(* IEC 61131-3 sources: SRCI_CLIENT_PLC/RobotLibrary/Library/POUs/General/MC_RobotTask (part 5) *)

           // Create log entry
           CreateLogMessagePara3 ( Timestamp   := SystemTime,
                                   MessageType := MessageType.CMD,
                                   Severity    := Severity.DEBUG,
                                   MessageCode := 0,
                                   MessageText := 'SyncWorkArea: Synchronization of WorkArea[{1}] triggered by PLC, SyncMode = {2}, SyncTime = {3}, SyncDirection = RC -> PLC',
                                   Para1       :=  DINT_TO_STRING(_rSyncIdx),
                                   Para2       :=  SYNC_MODE_TO_STRING(AxesGroup.Parameter.Plc.Parameter.SynchronizationModes.WorkAreas[SyncTime.AFTER_START_UP]),
                                   Para3       :=  SYNC_TIME_TO_STRING(SyncTime.AFTER_START_UP));
                                   RETURN;
         END_IF

         // Conflict triggered by RC ?
         IF ( NOT AxesGroup.State.SyncStateRc.InSync.WorkArea )
         THEN
           // get changed index
          _rSyncIdx := LIMIT(0, AxesGroup.State.SyncStateRc.UnSyncNo.WorkArea, AxesGroup.State.UnifiedWorkAreaIndex);
           // set timeout
           SetTimeout(PT := _rTimeout, rTimer := _rTimer);
           // inc step counter
          _rStep := 20; // -> read RC data and write it to PLC

           // Create log entry
           CreateLogMessagePara3 ( Timestamp   := SystemTime,
                                   MessageType := MessageType.CMD,
                                   Severity    := Severity.DEBUG,
                                   MessageCode := 0,
                                   MessageText := 'SyncWorkArea: Synchronization of WorkArea[{1}] triggered by RC, SyncMode = {2}, SyncTime = {3}, SyncDirection = RC -> PLC',
                                   Para1       :=  DINT_TO_STRING(_rSyncIdx),
                                   Para2       :=  SYNC_MODE_TO_STRING(AxesGroup.Parameter.Plc.Parameter.SynchronizationModes.WorkAreas[SyncTime.AFTER_START_UP]),
                                   Para3       :=  SYNC_TIME_TO_STRING(SyncTime.AFTER_START_UP));
                                   RETURN;
  			 END_IF

         // set timeout
         SetTimeout(PT := _rTimeout, rTimer := _rTimer);
         // jump back
        _rStep := 10;

    // ------------------------------------------
    // SyncMode : AUTOMATIC
    // ------------------------------------------
    13 : // Conflict triggerd by PLC ?
         IF ( NOT AxesGroup.State.SyncStatePlc.InSync.WorkArea )
         THEN
           // search for changed index
           FOR _rSyncIdx := 0 TO AxesGroup.State.UnifiedWorkAreaIndex
           DO
             IF ( AxesGroup.State.DataChanged.WorkArea[_rSyncIdx] )
             THEN
               // set timeout
               SetTimeout(PT := _rTimeout, rTimer := _rTimer);
               // inc step counter
              _rStep := 30; // -> write PLC data to RC
               EXIT;
  					 END_IF
           END_FOR

           // Create log entry
           CreateLogMessagePara3 ( Timestamp   := SystemTime,
                                   MessageType := MessageType.CMD,
                                   Severity    := Severity.DEBUG,
                                   MessageCode := 0,
                                   MessageText := 'SyncWorkArea: Synchronization of WorkArea[{1}] triggered by PLC, SyncMode = {2}, SyncTime = {3}, SyncDirection = PLC -> RC',
                                   Para1       :=  DINT_TO_STRING(_rSyncIdx),
                                   Para2       :=  SYNC_MODE_TO_STRING(AxesGroup.Parameter.Plc.Parameter.SynchronizationModes.WorkAreas[SyncTime.AFTER_START_UP]),
                                   Para3       :=  SYNC_TIME_TO_STRING(SyncTime.AFTER_START_UP));
                                   RETURN;
         END_IF

         // Conflict triggered by RC ?
         IF ( NOT AxesGroup.State.SyncStateRc.InSync.WorkArea )
         THEN
           // get changed index
          _rSyncIdx := LIMIT(0, AxesGroup.State.SyncStateRc.UnSyncNo.WorkArea, AxesGroup.State.UnifiedWorkAreaIndex);
           // set timeout
           SetTimeout(PT := _rTimeout, rTimer := _rTimer);
           // inc step counter
          _rStep := 20; // -> read RC data an write it to PLC

           // Create log entry
           CreateLogMessagePara3 ( Timestamp   := SystemTime,
                                   MessageType := MessageType.CMD,
                                   Severity    := Severity.DEBUG,
                                   MessageCode := 0,
                                   MessageText := 'SyncWorkArea: Synchronization of WorkArea[{1}] triggered by RC, SyncMode = {2}, SyncTime = {3}, SyncDirection = RC -> PLC',
                                   Para1       :=  DINT_TO_STRING(_rSyncIdx),
                                   Para2       :=  SYNC_MODE_TO_STRING(AxesGroup.Parameter.Plc.Parameter.SynchronizationModes.WorkAreas[SyncTime.AFTER_START_UP]),
                                   Para3       :=  SYNC_TIME_TO_STRING(SyncTime.AFTER_START_UP));
                                   RETURN;
  			 END_IF

         // set timeout
         SetTimeout(PT := _rTimeout, rTimer := _rTimer);
         // jump back
        _rStep := 10; // ST-FIX F95: was commented out

    // ------------------------------------------
    // Read Data from RC and write it to PLC
    // ------------------------------------------
    20 : IF (( NOT _readWorkArea.Busy  ) AND
             ( NOT _readWorkArea.Error ))
         THEN
           // set command parameter
          _readWorkArea.ParCmd.WorkAreaNo := _rSyncIdx;
           // execute command
          _readWorkArea.Execute := TRUE;
           // set timeout
           SetTimeout(PT := _rTimeout, rTimer := _rTimer);
           // inc step counter
          _rStep := _rStep + 1;
         ELSE
           // check error ?
           IF (_readWorkArea.Error)
           THEN
             ErrorID     := _readWorkArea.ErrorID;
             ErrorAddTxt := _readWorkArea.ErrorAddTxt;
           END_IF

           // timeout exceeded ?
           IF (CheckTimeout(_rTimer) = RobotLibraryConstants.OK)
           THEN
             ErrorID     := RobotLibraryErrorIdEnum.ERR_TIMEOUT_CMD;
             ErrorAddTxt := CONCAT(_stepName, DINT_TO_STRING(_rStep));
           END_IF
         END_IF

    21 : IF (( NOT _readWorkArea.Busy  ) AND
             ( NOT _readWorkArea.Error ) AND
             (     _readWorkArea.Done  ))
         THEN
           // reset execution
          _readWorkArea.Execute := FALSE;
           // ST-FIX F107: AUTOMATIC - the PLC data were changed while the RC data were read: the PLC
           // change is the most recent one and is written to the RC instead of being overwritten
           IF ( AxesGroup.Parameter.Plc.Parameter.SynchronizationModes.WorkAreas[SyncTime.AFTER_START_UP] = SyncMode.AUTOMATIC ) AND
              ( NOT IsWorkAreaEqual( Data1 := WorkAreas[_rSyncIdx].Data, Data2 := _workAreas[_rSyncIdx].Data, IgnoreTimestamp := TRUE ))
           THEN
             // set timeout
             SetTimeout(PT := _rTimeout, rTimer := _rTimer);
             // -> write PLC data to RC
            _rStep := 30;
             RETURN;
           END_IF
           // update internal WorkArea data
           WorkAreas[_rSyncIdx].Data := _readWorkArea.OutCmd.WorkAreaData;
          _workAreas[_rSyncIdx].Data := _readWorkArea.OutCmd.WorkAreaData;
           // set available bit
           WorkAreas[_rSyncIdx].Available := TRUE;
          _workAreas[_rSyncIdx].Available := TRUE;
           // set timeout
           SetTimeout(PT := _rTimeout, rTimer := _rTimer);
           // inc step counter
          // ST-FIX F20: write the RC data back to reset DataChanged on the RC (spec 5.6.7.4.2)
          IF ( AxesGroup.State.RobotData.RCSupportedFunctions.WriteWorkArea )
          THEN
            _rStep := 30;
          ELSE
            _rStep := 10;
          END_IF // -> jump to after startup
         ELSE
           // check error ?
           IF (_readWorkArea.Error)
           THEN
             ErrorID     := _readWorkArea.ErrorID;
             ErrorAddTxt := _readWorkArea.ErrorAddTxt;
             // reset available bit
             WorkAreas[_rSyncIdx].Available := FALSE;
            _workAreas[_rSyncIdx].Available := FALSE;
           END_IF

           // timeout exceeded ?
           IF (CheckTimeout(_rTimer) = RobotLibraryConstants.OK)
           THEN
             ErrorID     := RobotLibraryErrorIdEnum.ERR_TIMEOUT_CMD;
             ErrorAddTxt := CONCAT(_stepName, DINT_TO_STRING(_rStep));
           END_IF
         END_IF

    // ------------------------------------------
    // Write data from PLC to RC
    // ------------------------------------------
    30 : IF (( NOT _writeWorkArea.Busy  ) AND
             ( NOT _writeWorkArea.Error ))
         THEN
           // set command parameter
          _writeWorkArea.ParCmd.WorkAreaNo   := _rSyncIdx;
          _writeWorkArea.ParCmd.WorkAreaData :=  WorkAreas[_rSyncIdx].Data;
           // execute command
          _writeWorkArea.Execute := TRUE;
           // set timeout
           SetTimeout(PT := _rTimeout, rTimer := _rTimer);
           // inc step counter
          _rStep := _rStep + 1;
         ELSE
           // check error ?
           IF (_writeWorkArea.Error)
           THEN
             ErrorID     := _writeWorkArea.ErrorID;
             ErrorAddTxt := _writeWorkArea.ErrorAddTxt;;
           END_IF

           // timeout exceeded ?
           IF (CheckTimeout(_rTimer) = RobotLibraryConstants.OK)
           THEN
             ErrorID     := RobotLibraryErrorIdEnum.ERR_TIMEOUT_CMD;
             ErrorAddTxt := CONCAT(_stepName, DINT_TO_STRING(_rStep));
           END_IF
         END_IF

    31 : IF (( NOT _writeWorkArea.Busy  ) AND
             ( NOT _writeWorkArea.Error ) AND
             (     _writeWorkArea.Done  ))
         THEN
           // execute command
          _writeWorkArea.Execute := FALSE;
           // update internal WorkArea data
          _workAreas[_rSyncIdx] := WorkAreas[_rSyncIdx];
           // set available bit
           WorkAreas[_rSyncIdx].Available := TRUE;
          _workAreas[_rSyncIdx].Available := TRUE;
           // set timeout
           SetTimeout(PT := _rTimeout, rTimer := _rTimer);
           // inc step counter
          _rStep := 10; // -> jump to after startup;
         ELSE
           // check error ?
           IF (_writeWorkArea.Error)
           THEN
             SetWarning( WarningID := RobotLibraryWarningIdEnum.WARN_WORK_AREA_SYNC_FAILED_BY_ERROR_OF_READ_OR_WRITE_CMD, Overwrite :=  TRUE);
             // reset available bit
             WorkAreas[_rSyncIdx].Available := FALSE;
            _workAreas[_rSyncIdx].Available := FALSE;
           END_IF

           // timeout exceeded ?
           IF (CheckTimeout(_rTimer) = RobotLibraryConstants.OK)
           THEN
             ErrorID     := RobotLibraryErrorIdEnum.ERR_TIMEOUT_CMD;
             ErrorAddTxt := CONCAT(_stepName, DINT_TO_STRING(_rStep));
           END_IF
         END_IF

  ELSE
    // invalid step
    ErrorID     := RobotLibraryErrorIdEnum.ERR_INVALID_STEP;
    ErrorAddTxt := CONCAT(_stepName , DINT_TO_STRING(_stepCmd));
  END_CASE

END_METHOD

METHOD PRIVATE HandleTelegramStateCtrl
VAR_INPUT
END_VAR

  // Telegram Control
  // ----------------
  IF ( _lastTelegramControl <> GetHalfeByteLo(Telegram.PlcToRob.Header.AxesGroupID_Control))
  THEN
    // Create log entry
    CreateLogMessagePara2 ( Timestamp   := SystemTime,
                            MessageType := MessageType.CMD,
                            Severity    := Severity.INFO,
                            MessageCode := 0,
                            MessageText := 'SRCI Interface control changed from {1} to {2}',
                            Para1       := TELEGRAM_CONTROL_TO_STRING(_lastTelegramControl),
                            Para2       := TELEGRAM_CONTROL_TO_STRING(GetHalfeByteLo(Telegram.PlcToRob.Header.AxesGroupID_Control)));

    _lastTelegramControl := GetHalfeByteLo(Telegram.PlcToRob.Header.AxesGroupID_Control);
  END_IF

  // Telegram State
  // ----------------
  IF ( _lastTelegramState <> Telegram.RobToPlc.Header.TelegramState)
  THEN
    // Create log entry
    CreateLogMessagePara2 ( Timestamp   := SystemTime,
                            MessageType := MessageType.CMD,
                            Severity    := Severity.INFO,
                            MessageCode := 0,
                            MessageText := 'SRCI Interface state changed from {1} to {2}',
                            Para1       := TELEGRAM_STATE_TO_STRING(_lastTelegramState),
                            Para2       := TELEGRAM_STATE_TO_STRING(Telegram.RobToPlc.Header.TelegramState));

    // Check Interface changed after being initialized ?
    IF ((  Enable                                                                          ) AND
        ( _lastTelegramState                      = TelegramState.INITIALIZED              ) AND
       ((  Telegram.RobToPlc.Header.TelegramState = TelegramState.READY_FOR_INITIALIZATION ) OR
        (  Telegram.RobToPlc.Header.TelegramState = TelegramState.READY_TO_RESUME          )))
    THEN
      // the error 16#80A7 (interface reset after the initialization) is set in OnCall (ST-FIX F65)
      ;
  	END_IF

    // apply new telegram state
   _lastTelegramState := Telegram.RobToPlc.Header.TelegramState;
  END_IF

END_METHOD

METHOD HandleUserData
VAR_IN_OUT
   /// Robot assignment of function
  AxesGroup    : AxesGroup;
  ///  User data stored on the PLC according to Table 6-10
  UserData     : UserData;
END_VAR

  // Common
  UserData.LogLevel                          := LogLevel;

  UserData.PLCManufacturedID                 := _parCfg.Plc.Parameter.ManufacturedID;
  UserData.PLCOrderID                        := _parCfg.Plc.Parameter.OrderID;
  UserData.PLCSerialNumber                   := _parCfg.Plc.Parameter.SerialNumber;
  UserData.PLCFirmwareVersion                := _parCfg.Plc.Parameter.FirmwareVersion;
  UserData.PLCInterfaceVersion               := _parCfg.Plc.Parameter.InterfaceVersion;
  UserData.PLCLibraryVersion                 :=  RobotLibraryConstants.PLCLibraryVersion;

  // Communication
  UserData.LifeSignTimeOut                   := _parCfg.Com.LifeSignTimeOut;

  // Plc Parameter
  UserData.SynchronizationModes              := _parCfg.Plc.Parameter.SynchronizationModes;
  UserData.EnableSync                        :=  SyncModesToDataEnableSync(Value := _parCfg.Plc.Parameter.SynchronizationModes);

  // Robot Parameter
  UserData.DelayTime                         := _parCfg.Rob.Parameter.DelayTime;
  UserData.WaitForNrOfCmd                    := _parCfg.Rob.Parameter.WaitForNrOfCmd;
  UserData.WaitAtBlendingZone                := _parCfg.Rob.Parameter.WaitAtBlendingZone;
  UserData.AllowSecSeqWhileSubprogram        := _parCfg.Rob.Parameter.AllowSecSeqWhileSubprogram;
  UserData.AllowDynamicBlending              := _parCfg.Rob.Parameter.AllowDynamicBlending;
  UserData.SyncReaction                      := _parCfg.Rob.Parameter.SyncReaction;
  UserData.SyncDelay                         := _parCfg.Rob.Parameter.SyncDelay;
  UserData.MessageLevel                      := _parcfg.Rob.Parameter.MessageLevel;

  // ReadRobotData
  UserData.RCManufacturer                    := AxesGroup.State.RobotData.RCManufacturer;
  UserData.RCOrderID                         := AxesGroup.State.RobotData.RCOrderID;
  UserData.RCSerialNumber                    := AxesGroup.State.RobotData.RCSerialNumber;
  UserData.RASerialNumber                    := AxesGroup.State.RobotData.RASerialNumber;
  UserData.RCFirmwareVersion                 := AxesGroup.State.RobotData.RCFirmwareVersion;

  UserData.RCInterpreterVersion := AxesGroup.State.RobotData.RCInterpreterVersionNumber; // ST-FIX F163: was characters 1/2/3 of the text

  UserData.AxisJointUsed                     := AxesGroup.State.RobotData.AxisJointUsed;
  UserData.AxisExternalUsed                  := AxesGroup.State.RobotData.AxisExternalUsed;
  UserData.AxisJointUnit                     := AxesGroup.State.RobotData.AxisJointUnit;
  UserData.AxisExternalUnit                  := AxesGroup.State.RobotData.AxisExternalUnit;
  UserData.RCSupportedFunctions              := AxesGroup.State.RobotData.RCSupportedFunctions;

  UserData.BrakeTestRequired                 := AxesGroup.State.ConfigurationData.BrakeTestRequired;
  UserData.PathAccuracyMode                  := AxesGroup.State.ConfigurationData.PathAccuracyMode;
  UserData.AvoidSingularity                  := AxesGroup.State.ConfigurationData.AvoidSingularity;
  UserData.ConstantVelocitySupported         := AxesGroup.State.ConfigurationData.ConstantVelocitySupported;
  UserData.StepModeExactStopActive           := AxesGroup.State.ConfigurationData.StepModeExactStopActive;
  UserData.StepModeBlendingActive            := AxesGroup.State.ConfigurationData.StepModeBlendingActive;
  UserData.AcceleratingSupported             := AxesGroup.State.ConfigurationData.AcceleratingSupported;
  UserData.DeceleratingSupported             := AxesGroup.State.ConfigurationData.DecceleratingSupported;

  UserData.Initialized                       := Initialized;
  UserData.Synchronized                      := Synchronized;

  // Cyclic data
  UserData.RCSRCIVersion                     := AxesGroup.Cyclic.RobToPlc.SRCIVersion;
  UserData.IsMoving                          := AxesGroup.Cyclic.RobToPlc.StatusRobotArm.IsMoving;
  UserData.PrimarySequencePaused             := AxesGroup.Cyclic.RobToPlc.StatusRobotArm.PrimarySequencePaused;
  UserData.InPrimaryPos                      := AxesGroup.Cyclic.RobToPlc.StatusRobotArm.InPrimaryPos;
  UserData.SecondarySequenceActive           := AxesGroup.Cyclic.RobToPlc.StatusRobotArm.SecondarySequenceActive;
  UserData.ErrorPending                      := AxesGroup.Cyclic.RobToPlc.StatusRobotArm.ErrorPending;
  UserData.RestartInProgress                 := AxesGroup.Cyclic.RobToPlc.StatusRobotArm.RestartInProgress;
  UserData.Enabled                           := AxesGroup.Cyclic.RobToPlc.StatusRobotArm.Enabled;
  UserData.Idle                              := AxesGroup.Cyclic.RobToPlc.StatusRobotArm.RaSequenceState = RaSequenceState.IDLE;
  UserData.Executing                         := AxesGroup.Cyclic.RobToPlc.StatusRobotArm.RaSequenceState = RaSequenceState.EXECUTING;
  UserData.Interrupted                       := AxesGroup.Cyclic.RobToPlc.StatusRobotArm.RaSequenceState = RaSequenceState.INTERRUPTED;
  UserData.IsBlending                        := AxesGroup.Cyclic.RobToPlc.StatusRobotArm.IsBlending;
  UserData.OperationMode                     := AxesGroup.Cyclic.RobToPlc.StatusRobotArm.OperationMode;
  UserData.CollisionDetectionEnabled         := AxesGroup.Parameter.Rob.Parameter.CollisionDetectionEnabled; // ST-FIX F169: the status word bit is always FALSE
  UserData.CollisionDetected                 := AxesGroup.Cyclic.RobToPlc.StatusRobotArm.CollisionDetected;
  UserData.RestartRequested                  := AxesGroup.Cyclic.RobToPlc.StatusRobotArm.RestartRequested;
  UserData.Accelerating                      := AxesGroup.Cyclic.RobToPlc.StatusRobotArm.Accelerating;
  UserData.Decelerating                      := AxesGroup.Cyclic.RobToPlc.StatusRobotArm.Decelerating;
  UserData.ConstantVelocity                  := AxesGroup.Cyclic.RobToPlc.StatusRobotArm.ConstantVelocity;
  UserData.ActualOverride                    := PERCENT_UINT_TO_REAL( Value := AxesGroup.Cyclic.RobToPlc.Override, IsOptional := FALSE);

  // Cyclic optional data
  UserData.CartesianPosition                 := AxesGroup.CyclicOptional.RobToPlc.CartesianPosition;
  UserData.ExtCartesianPosition              := AxesGroup.CyclicOptional.RobToPlc.CartesianPositionExt;
  UserData.JointPosition                     := AxesGroup.CyclicOptional.RobToPlc.JointPosition;
  UserData.ExtJointPosition                  := AxesGroup.CyclicOptional.RobToPlc.JointPositionExt;

  // Synchronizing
  UserData.ToolDataSynchronizing             := AxesGroup.State.Synchronizing.Tool;
  UserData.FrameDataSynchronizing            := AxesGroup.State.Synchronizing.Frame;
  UserData.LoadDataSynchronizing             := AxesGroup.State.Synchronizing.Load;
  UserData.WorkAreaDataSynchronizing         := AxesGroup.State.Synchronizing.WorkAreas;
  UserData.SWLimitsSynchronizing             := AxesGroup.State.Synchronizing.SwLimits;
  UserData.DefaultDynamicsSynchronizing      := AxesGroup.State.Synchronizing.DefaultDynamics;
  UserData.ReferenceDynamicsSynchronizing    := AxesGroup.State.Synchronizing.ReferenceDynamics;

  UserData.ActivateTwoSequences              := _parCfg.Com.TwoSequences;
  UserData.ReadingCartesianPosition          :=  AxesGroup.State.ReadingCartesianPosition;
  UserData.ReadingExtCartesianPosition       :=  AxesGroup.State.ReadingCartesianPositionExt;
  UserData.ReadingJointPosition              :=  AxesGroup.State.ReadingJointPosition;
  UserData.ReadingExtJointPosition           :=  AxesGroup.State.ReadingJointPositionExt;

END_METHOD

PROPERTY PROTECTED HasError : Bool

GET
VAR
END_VAR

  HasError := ErrorID <> RobotLibraryErrorIdEnum.NO_ERROR;

END_GET

PROPERTY PROTECTED HasInfo : BOOL

GET
VAR
END_VAR

  HasInfo := InfoID <> RobotLibraryInfoIdEnum.NO_INFO;

END_GET

PROPERTY PROTECTED HasWarning : BOOL

GET
VAR
END_VAR

  HasWarning := WarningID <> RobotLibraryWarningIdEnum.NO_WARNING;

END_GET

METHOD PRIVATE OnCall
VAR_IN_OUT
   /// Robot assignment of function
  AxesGroup : AxesGroup;
END_VAR

  // map numeric value to enum, so that the corresponding message text is directly shown by the tooltip
  ErrorIdEnum   := ErrorId;
  WarningIdEnum := WarningId;
  InfoIdEnum    := InfoId;

  Error := HasError;

  // Check Payload and In/Out data size
  IF (( ROBOT_IN_DATA_SIZE  < 64 ) OR
      ( ROBOT_OUT_DATA_SIZE < 64 ))
  THEN
    SetError(ErrorID := RobotLibraryErrorIdEnum.ERR_INVALID_LIBRARY_PARA, Overwrite := TRUE );
    RETURN;
  END_IF

  // Check AxesGroupID valid
  IF (( AxesGroupID < RobotLibraryConstants.AXES_GROUP_ID_MIN ) OR
      ( AxesGroupID > RobotLibraryConstants.AXES_GROUP_ID_MAX ))
  THEN
    // ST-FIX F138: client error of the specification (16#80AA, table 7-2) instead of the internal ID 3
    SetError( ErrorID := RobotLibraryErrorIdEnum.ERR_AXESGROUP_ID_INVALID_0x80AA, Overwrite := TRUE );
    RETURN;
  END_IF

  // Reset flag for initialization / Synchronization
  IF ( Initialized OR Synchronized) AND ( AxesGroup.Cyclic.RobToPlc.TelegramState <> TelegramState.INITIALIZED)
  THEN
    // Reset initialized flag
    Initialized := FALSE;
    // Reset Synchronized flag
    Synchronized := FALSE;
    // Set error
    // ST-FIX F65: reason of the loss of the initialization (table 7-2): RI error of the RC in the
    // telegram state (16#A1..16#AD), interface reset by the RC (16#80A7) or unknown (16#80A2)
    IF (( AxesGroup.Cyclic.RobToPlc.TelegramState >= TelegramState.ERROR_161_TELEGRAM_CONTROL_MISMATCH_TELEGRAM_STATE ) AND
        ( AxesGroup.Cyclic.RobToPlc.TelegramState <= TelegramState.ERROR_173_SERVER_CONNECTION_LOST                   ))
    THEN
      SetError( ErrorID := AxesGroup.Cyclic.RobToPlc.TelegramState, Overwrite := TRUE );
      // Create log entry
      CreateLogMessagePara1 ( Timestamp   := SystemTime,
                              MessageType := MessageType.CMD,
                              Severity    := Severity.ERROR,
                              MessageCode := ErrorID,
                              MessageText := 'Initialization lost: RI error {1} of the RC',
                              Para1       := TELEGRAM_STATE_TO_STRING(AxesGroup.Cyclic.RobToPlc.TelegramState));
    ELSIF (( AxesGroup.Cyclic.RobToPlc.TelegramState = TelegramState.READY_FOR_INITIALIZATION ) OR
           ( AxesGroup.Cyclic.RobToPlc.TelegramState = TelegramState.READY_TO_RESUME          ))
    THEN
      SetError( ErrorID := RobotLibraryErrorIdEnum.ERR_INTERFACE_WAS_RESET_AFTER_INIT_0x80A7, Overwrite := TRUE );
      // Create log entry
      CreateLogMessagePara1 ( Timestamp   := SystemTime,
                              MessageType := MessageType.CMD,
                              Severity    := Severity.ERROR,
                              MessageCode := ErrorID,
                              MessageText := 'Initialization lost: interface was reset by the RC (state {1})',
                              Para1       := TELEGRAM_STATE_TO_STRING(AxesGroup.Cyclic.RobToPlc.TelegramState));
    ELSE
      SetError( ErrorID := RobotLibraryErrorIdEnum.ERR_INIT_LOST_UNKNOWN_0x80A2, Overwrite := TRUE );
      // Create log entry
      CreateLogMessagePara1 ( Timestamp   := SystemTime,
                              MessageType := MessageType.CMD,
                              Severity    := Severity.ERROR,
                              MessageCode := ErrorID,
                              MessageText := 'Initialization lost: unknown reason (state {1})',
                              Para1       := TELEGRAM_STATE_TO_STRING(AxesGroup.Cyclic.RobToPlc.TelegramState));
    END_IF
  END_IF

  // Warning for ACR Registers running low
  IF ( AxesGroup.Acyclic.ActiveCommandRegister.CurrentAcrUsagePercent > RobotLibraryParameter.ACR_USAGE_WARNING_LIMIT )
  THEN
    SetWarning( WarningID := RobotLibraryWarningIdEnum.WARN_ACR_FREE_ENTRIES_LOW, Overwrite := TRUE);
  END_IF

  // Check ToolData boundary
  IF ( AxesGroup.SystemData.ToolDataMin  <> 0 )
  THEN
    SetWarning( WarningID := RobotLibraryWarningIdEnum.WARN_TOOL_DATA_ARRAY_NOT_START_AT_ZERO, Overwrite := FALSE );
  END_IF

  // Check FrameData boundary
  IF ( AxesGroup.SystemData.FrameDataMin <> 0 ) AND ( NOT HasWarning )
  THEN
    SetWarning( WarningID := RobotLibraryWarningIdEnum.WARN_FRAME_DATA_ARRAY_NOT_START_AT_ZERO, Overwrite := FALSE );
  END_IF

  // Check WorkAreas boundary
  IF ( AxesGroup.SystemData.WorkAreasMin <> 0 ) AND ( NOT HasWarning )
  THEN
    SetWarning( WarningID := RobotLibraryWarningIdEnum.WARN_FRAME_DATA_ARRAY_NOT_START_AT_ZERO, Overwrite := FALSE);
  END_IF

  // Check configuration parameter changed ?
  CheckParameterChanged(AxesGroup := AxesGroup);

END_METHOD

METHOD OnExecRun : DINT
VAR_IN_OUT
  /// Robot assignment of function
  AxesGroup         : AxesGroup;
END_VAR

  // building rising and falling edges
  _enable_R( CLK := Enable);
  _enable_F( CLK := Enable);

  IF ( _enable_F.Q)
  THEN
    Reset(AxesGroup := AxesGroup);
  END_IF

  OnExecRun := RobotLibraryConstants.RUNNING;

  CASE _stepCmd OF

    00:  IF ( _enable_R.Q )
         THEN
           // Create log entry
           CreateLogMessage ( Timestamp   := SystemTime,
                              MessageType := MessageType.CMD,
                              Severity    := Severity.INFO,
                              MessageCode := 0,
                              MessageText := 'Robot Task Enabled');

           // reset the rising edge
          _enable_R();
           // set busy flag
           Busy := TRUE;
           // set timeout
           SetTimeout(PT := _timeoutCmd, rTimer := _timerCmd);
           // Reset FastStop
           AxesGroup.Cyclic.PlcToRob.FastStop := 0;
           // Reset Active command register
           AxesGroup.Acyclic.ActiveCommandRegister.Reset();
           // ST-FIX F23: the RC is still initialized from the previous enable (ACR, SEQ/ACK)
           // -> reset the interface on the RC as well
           _restartReset := AxesGroup.Cyclic.RobToPlc.TelegramState = TelegramState.INITIALIZED;
           IF ( _restartReset )
           THEN
             AxesGroup.Cyclic.PlcToRob.Control := ControlHalfByte.RESET;
           END_IF

           // check parameter valid
           IF ( CheckParameterValid(AxesGroup := AxesGroup) )
           THEN
             // take configuration parameter if not yet enabled
            _parCfg := ParCfg;
            // ST-FIX F103: number of telegram sequences of this configuration (not of the previous enable)
            IF ( _parCfg.Com.TwoSequences )
            THEN
              AxesGroup.State.SequenceCountSend := 1;
            ELSE
              AxesGroup.State.SequenceCountSend := 0;
            END_IF
            // ST-FIX F79: no error state of the RC seen yet in this initialization
            _initErrorState := TelegramState.UNDEFINED;
             // inc step counter
            _stepCmd := _stepCmd + 1;
           END_IF
         END_IF

    01:  // ST-FIX F153: INITIALIZED without a request of this RobotTask: the RC is still
  // initialized from an earlier connection -> reset the interface on the RC first
  IF (( AxesGroup.Cyclic.RobToPlc.TelegramState = TelegramState.INITIALIZED ) AND
      ( AxesGroup.Cyclic.PlcToRob.Control       = ControlHalfByte.NONE      ) AND
      ( NOT _restartReset                                                   ))
  THEN
    AxesGroup.Cyclic.PlcToRob.Control := ControlHalfByte.RESET;
    _restartReset := TRUE;
  END_IF

  // ST-FIX F23: wait until the RC left the state INITIALIZED of the previous enable
  IF ( _restartReset )
  THEN
    IF ( AxesGroup.Cyclic.RobToPlc.TelegramState <> TelegramState.INITIALIZED )
    THEN
      _restartReset := FALSE;
    END_IF
  ELSE
  CASE AxesGroup.Cyclic.RobToPlc.TelegramState  OF

           TelegramState.UNDEFINED : ;

           TelegramState.ERROR_161_TELEGRAM_CONTROL_MISMATCH_TELEGRAM_STATE..TelegramState.ERROR_172_TELEGRAM_NUMBER_NOT_SUPPORTED:

             // ST-FIX F79: remember the error state for the init timeout
             _initErrorState := AxesGroup.Cyclic.RobToPlc.TelegramState;

             // clear error
             AxesGroup.Cyclic.PlcToRob.Control := ControlHalfByte.ACK_ERROR;
             AxesGroup.Cyclic.PlcToRob.Control := ControlHalfByte.RESET; // always a reset, so that on the robot side the ACR is reseted

           TelegramState.ERROR_173_SERVER_CONNECTION_LOST:

             // Reset interface including the ACR register on server side
             AxesGroup.Cyclic.PlcToRob.Control := ControlHalfByte.RESET;

           TelegramState.READY_TO_RESUME :

             // Resume
             AxesGroup.Cyclic.PlcToRob.Control := ControlHalfByte.RESUME;

           TelegramState.READY_FOR_INITIALIZATION:

             // Request initialization
             AxesGroup.Cyclic.PlcToRob.Control := ControlHalfByte.INITIALIZE;

           TelegramState.INITIALIZED:

             // Reset Telegram Control
             AxesGroup.Cyclic.PlcToRob.Control := ControlHalfByte.NONE;

             // Check SRCI Version is compatible ?
             IF ( AxesGroup.Cyclic.RobToPlc.SRCIVersion.MajorVersion = RobotLibraryConstants.SRCIVersion.MajorVersion )
             THEN
               // set timeout
               SetTimeout(PT := _timeoutCmd, rTimer := _timerCmd);
               // inc step counter
              _stepCmd := _stepCmd + 1;
             ELSE
               // set error
               ErrorID     := RobotLibraryErrorIdEnum.ERR_SRCI_MAJOR_VERSION_INCOMPATIBLE_0x80A4;
               ErrorAddTxt := CONCAT('_stepCmd = ' , DINT_TO_STRING(_stepCmd));
             END_IF

         ELSE
           // TelegrammState in error
           SetError( ErrorID := RobotLibraryErrorIdEnum.ERR_INIT_LOST_UNKNOWN_0x80A2, Overwrite := TRUE ); // ST-FIX F65: unknown state (16#A2 is the RI error of the RC)
             // Create log entry
             CreateLogMessagePara1 ( Timestamp   := SystemTime,
                                     MessageType := MessageType.CMD,
                                     Severity    := Severity.ERROR,
                                     MessageCode := ErrorID,
                                     MessageText := 'Initialization lost: unknown telegram state {1}',
                                     Para1       := TELEGRAM_STATE_TO_STRING(AxesGroup.Cyclic.RobToPlc.TelegramState));
           ErrorAddTxt := CONCAT('_stepCmd = ' , DINT_TO_STRING(_stepCmd));
         END_CASE
  END_IF

         // timeout exceeded ?
         IF (CheckTimeout(_timerCmd) = RobotLibraryConstants.OK)
         THEN
           // Check Telegram State error ?
           IF (( AxesGroup.Cyclic.RobToPlc.TelegramState >= TelegramState.ERROR_161_TELEGRAM_CONTROL_MISMATCH_TELEGRAM_STATE ) AND // ST-FIX F15
               ( AxesGroup.Cyclic.RobToPlc.TelegramState <= TelegramState.ERROR_173_SERVER_CONNECTION_LOST                   ))
           THEN
             ErrorID     := AxesGroup.Cyclic.RobToPlc.TelegramState;
             ErrorAddTxt := CONCAT('_stepCmd = ' , DINT_TO_STRING(_stepCmd));
           ELSIF ( _initErrorState <> TelegramState.UNDEFINED ) // ST-FIX F79: error state seen during the initialization
           THEN
             ErrorID     := _initErrorState;
             ErrorAddTxt := CONCAT('_stepCmd = ' , DINT_TO_STRING(_stepCmd));
           ELSE
             ErrorID     := RobotLibraryErrorIdEnum.ERR_TIMEOUT_CMD;
             ErrorAddTxt := CONCAT('_stepCmd = ' , DINT_TO_STRING(_stepCmd));
           END_IF
         END_IF

    02: IF (( NOT _readMessages.Busy  ) AND
            ( NOT _readMessages.Error ))
        THEN
          // start function block
         _readMessages.Enable := TRUE;
         _readMessages.ParCmd.MsgID := 0;
         _readMessages.ParCmd.MessageLevel := _parCfg.Rob.Parameter.MessageLevel;

          // set timeout
          SetTimeout(PT := _timeoutCmd, rTimer := _timerCmd);
          // inc step counter
         _stepCmd := _stepCmd + 1;
        ELSE
          // check error ?
          IF (_readMessages.Error)
          THEN
            ErrorID     := _readMessages.ErrorID;
            ErrorAddTxt := _readMessages.ErrorAddTxt;;
          END_IF
          // timeout exceeded ?
          IF (CheckTimeout(_timerCmd) = RobotLibraryConstants.OK)
          THEN
            ErrorID     := RobotLibraryErrorIdEnum.ERR_TIMEOUT_CMD;
            ErrorAddTxt := CONCAT('_stepCmd = ' , DINT_TO_STRING(_stepCmd));
          END_IF
        END_IF

    03: IF ((     _readMessages.Enabled ) AND
            ( NOT _readMessages.Error   ))
        THEN
          // ---------------------------------------------------------------
          // !!! ReadMessages must stay active for the Message mechanism !!!
          // ---------------------------------------------------------------
          // ReadMessages.Enable := FALSE;
          // set timeout
          SetTimeout(PT := _timeoutCmd, rTimer := _timerCmd);
          // inc step counter
         _stepCmd := _stepCmd + 1;
        ELSE
           // check error ?
           IF (_readMessages.Error)
           THEN
             ErrorID     := _readMessages.ErrorID;
             ErrorAddTxt := _readMessages.ErrorAddTxt;;
           END_IF

           // timeout exceeded ?
           IF (CheckTimeout(_timerCmd) = RobotLibraryConstants.OK)
           THEN
             ErrorID     := RobotLibraryErrorIdEnum.ERR_TIMEOUT_CMD;
             ErrorAddTxt := CONCAT('_stepCmd = ' , DINT_TO_STRING(_stepCmd));
           END_IF
         END_IF

    04: IF (( NOT _exchangeConfiguration.Busy  ) AND
            ( NOT _exchangeConfiguration.Error ))
        THEN
          // set command parameter
         _exchangeConfiguration.ParCmd.LogLevel                           :=  LogLevel;
         _exchangeConfiguration.ParCmd.WaitAtBlendingZone                 := _parCfg.Rob.Parameter.WaitAtBlendingZone;
         _exchangeConfiguration.ParCmd.AllowSecSeqWhileSubprogram         := _parCfg.Rob.Parameter.AllowSecSeqWhileSubprogram;
         _exchangeConfiguration.ParCmd.AllowDynamicBlending               := _parCfg.Rob.Parameter.AllowDynamicBlending;
         _exchangeConfiguration.ParCmd.DelayTime                          := _parCfg.Rob.Parameter.DelayTime;
         _exchangeConfiguration.ParCmd.WaitForNrOfCmd                     := _parCfg.Rob.Parameter.WaitForNrOfCmd;
         _exchangeConfiguration.ParCmd.LifeSignTimeOut                    :=  TIME_TO_UINT(_parCfg.Com.LifeSignTimeOut);
         _exchangeConfiguration.ParCmd.SyncDelay                          := _parCfg.Rob.Parameter.SyncDelay;
         _exchangeConfiguration.ParCmd.SyncReaction                       := _parCfg.Rob.Parameter.SyncReaction;
         _exchangeConfiguration.ParCmd.DataEnableSync                     :=  SyncModesToDataEnableSync(Value := _parCfg.Plc.Parameter.SynchronizationModes);
         _exchangeConfiguration.ParCmd.DataInSync.ToolsInSync             :=  FALSE;
         _exchangeConfiguration.ParCmd.DataInSync.FramesInSync            :=  FALSE;
         _exchangeConfiguration.ParCmd.DataInSync.LoadsInSync             :=  FALSE;
         _exchangeConfiguration.ParCmd.DataInSync.WorkAreasInSync         :=  FALSE;
         _exchangeConfiguration.ParCmd.DataInSync.SoftwareLimitsInSync    :=  FALSE;
         _exchangeConfiguration.ParCmd.DataInSync.DefaultDynamicsInSync   :=  FALSE;
         _exchangeConfiguration.ParCmd.DataInSync.ReferenceDynamicsInSync :=  FALSE;

          // start function block
         _exchangeConfiguration.Enable := TRUE;
          // set timeout
          SetTimeout(PT := _timeoutCmd, rTimer := _timerCmd);
          // inc step counter
         _stepCmd := _stepCmd + 1;
        ELSE
          // check error ?
          IF (_exchangeConfiguration.Error)
          THEN
            ErrorID     := _exchangeConfiguration.ErrorID;
            ErrorAddTxt := _exchangeConfiguration.ErrorAddTxt;;
          END_IF

          // timeout exceeded ?
          IF (CheckTimeout(_timerCmd) = RobotLibraryConstants.OK)
          THEN
            ErrorID     := RobotLibraryErrorIdEnum.ERR_TIMEOUT_CMD;
            ErrorAddTxt := CONCAT('_stepCmd = ' , DINT_TO_STRING(_stepCmd));
          END_IF
        END_IF

    05: IF ((     _exchangeConfiguration.Enabled ) AND
            ( NOT _exchangeConfiguration.Error   ))
        THEN
          // ---------------------------------------------------------------------
          // !!! ExchangeConfiguration must stay active for the Sync mechanism !!!
          // ---------------------------------------------------------------------
          // ExchangeConfiguration.Enable := FALSE;
          // set timeout
          SetTimeout(PT := _timeoutCmd, rTimer := _timerCmd);
          // inc step counter
         _stepCmd := _stepCmd + 1;
        ELSE
          // check error ?
          IF (_exchangeConfiguration.Error)
          THEN
            ErrorID     := _exchangeConfiguration.ErrorID;
            ErrorAddTxt := _exchangeConfiguration.ErrorAddTxt;;
          END_IF

          // timeout exceeded ?
          IF (CheckTimeout(_timerCmd) = RobotLibraryConstants.OK)
          THEN
            ErrorID     := RobotLibraryErrorIdEnum.ERR_TIMEOUT_CMD;
            ErrorAddTxt := CONCAT('_stepCmd = ' , DINT_TO_STRING(_stepCmd));
          END_IF
        END_IF

    06: IF (( NOT _readRobotData.Busy  ) AND
            ( NOT _readRobotData.Error ))
        THEN
          // start function block
         _readRobotData.Execute := TRUE;
          // set timeout
          SetTimeout(PT := _timeoutCmd, rTimer := _timerCmd);
          // inc step counter
         _stepCmd := _stepCmd + 1;
        ELSE
          // check error ?
          IF (_readRobotData.Error)
          THEN
            ErrorID     := _readRobotData.ErrorID;
            ErrorAddTxt := _readRobotData.ErrorAddTxt;;
          END_IF
          // timeout exceeded ?
          IF (CheckTimeout(_timerCmd) = RobotLibraryConstants.OK)
          THEN
            ErrorID     := RobotLibraryErrorIdEnum.ERR_TIMEOUT_CMD;
            ErrorAddTxt := CONCAT('_stepCmd = ' , DINT_TO_STRING(_stepCmd));
          END_IF
        END_IF

    07: IF ((     _readRobotData.Done  ) AND
            ( NOT _readRobotData.Busy  ) AND
            ( NOT _readRobotData.Error ))
        THEN
          // set initialized flag
          Initialized := TRUE;
          // start function block
         _readRobotData.Execute := FALSE;
          // set timeout
          SetTimeout(PT := _timeoutCmd, rTimer := _timerCmd);
          // inc step counter
         _stepCmd := _stepCmd + 1;
         ELSE
           // check error ?
           IF (_readRobotData.Error)
           THEN
             ErrorID     := _readRobotData.ErrorID;
             ErrorAddTxt := _readRobotData.ErrorAddTxt;;
           END_IF

           // timeout exceeded ?
           IF (CheckTimeout(_timerCmd) = RobotLibraryConstants.OK)
           THEN
             ErrorID     := RobotLibraryErrorIdEnum.ERR_TIMEOUT_CMD;
             ErrorAddTxt := CONCAT('_stepCmd = ' , DINT_TO_STRING(_stepCmd));
           END_IF
         END_IF

    08:  // Update Initialized state
         // ST-FIX F131: Initialized stays TRUE while Synchronized (RI state "Synchronized" includes the
         // initialization); otherwise CheckParameterChanged did not run while synchronized
         Initialized := NOT Error;
         // ST-FIX F29: the next line overwrote the error check above
         // Initialized := NOT Synchronized;

         // Wait for task disable
         IF ( NOT Enable)
         THEN
           // Reset active command register
           AxesGroup.Acyclic.ActiveCommandRegister.Reset();
           // reset internal variables
           Reset(AxesGroup := AxesGroup);
           // Reset step counter
          _stepCmd := 0;
           // finished okay
           OnExecRun := RobotLibraryConstants.OK;
         END_IF

  ELSE
    // invalid step
    ErrorID     := RobotLibraryErrorIdEnum.ERR_INVALID_STEP;
    ErrorAddTxt := CONCAT('_stepCmd = ' , DINT_TO_STRING(_stepCmd));
  END_CASE

END_METHOD

METHOD PROTECTED ParseRecvPayload
VAR_IN_OUT
  /// Robot assignment of function
  AxesGroup   : AxesGroup;
  /// Inputs of PLC for communication from RC
  RobotInData : ARRAY[*] OF BYTE;
END_VAR

  // reset all variables and payload
  RecvData.Reset();
  // Call RecvData FB, update payload and size
  RecvData(Payload := RobotInData, PayloadSize := ROBOT_IN_DATA_SIZE);

  // check new data to receive ?
  // ST-FIX F140: also new data of the 2nd sequence
  IF ( Telegram.RobToPlc.Sequence[0].Header.SEQ_ACK <> AxesGroup.State.LastACK[0] ) OR
     ( Telegram.RobToPlc.Sequence[1].Header.SEQ_ACK <> AxesGroup.State.LastACK[1] )
  THEN
    // delete old telegram data
    SysDepMemSet(pDest := ADR(Telegram.RobToPlc), Value := 0 , DataLen := SIZEOF(Telegram.RobToPlc));
  END_IF

  ParseRecvPayloadHeader        ( AxesGroup := AxesGroup);
  ParseRecvPayloadCyclic        ( AxesGroup := AxesGroup);
  ParseRecvPayloadCyclicOptional( AxesGroup := AxesGroup);
  ParseRecvPayloadSequence      ( AxesGroup := AxesGroup);
  ParseRecvPayloadFooter        ( AxesGroup := AxesGroup);
  ParseRecvPayloadLogging       ( AxesGroup := AxesGroup);

  AxesGroup.State.LastACK[0] := Telegram.RobToPlc.Sequence[0].Header.SEQ_ACK;
  AxesGroup.State.LastACK[1] := Telegram.RobToPlc.Sequence[1].Header.SEQ_ACK;

END_METHOD

METHOD PROTECTED ParseRecvPayloadCyclic
VAR_IN_OUT
  /// Robot assignment of function
  AxesGroup: AxesGroup;
END_VAR

END_METHOD

METHOD PROTECTED ParseRecvPayloadCyclicOptional
VAR_IN_OUT
  /// Robot assignment of function
  AxesGroup    : AxesGroup;
END_VAR

VAR
  /// internal index for loops
 _idx : DINT;
END_VAR

  // AxesGroup.OptionalCyclic.RobToPlc.SubProgramData {{{
  IF ( AxesGroup.CyclicOptional.RobToPlc.SubProgramData.Active )
  THEN
    FOR _idx := 0 TO  RobotLibraryConstants.CYCLIC_SUB_PROGRAM_DATA_MAX (* ST-FIX F179 *)
    DO
      Telegram.RobToPlc.CyclicOptional.SubProgramData.Data[_idx] := RecvData.GetByte();
    END_FOR
  END_IF
  // }}}

  // AxesGroup.OptionalCyclic.RobToPlc.CartesianPos {{{
  IF ( AxesGroup.CyclicOptional.RobToPlc.CartesianPosition.Active )
  THEN
    Telegram.RobToPlc.CyclicOptional.CartesianPosition.X                    := RecvData.GetReal();
    Telegram.RobToPlc.CyclicOptional.CartesianPosition.Y                    := RecvData.GetReal();
    Telegram.RobToPlc.CyclicOptional.CartesianPosition.Z                    := RecvData.GetReal();
    Telegram.RobToPlc.CyclicOptional.CartesianPosition.Rx                   := RecvData.GetReal();
    Telegram.RobToPlc.CyclicOptional.CartesianPosition.Ry                   := RecvData.GetReal();
    Telegram.RobToPlc.CyclicOptional.CartesianPosition.Rz                   := RecvData.GetReal();
    Telegram.RobToPlc.CyclicOptional.CartesianPosition.Config               := RecvData.GetWord();
    Telegram.RobToPlc.CyclicOptional.CartesianPosition.Turns_J2_J1          := RecvData.GetByte();
    Telegram.RobToPlc.CyclicOptional.CartesianPosition.Turns_J4_J3          := RecvData.GetByte();
    Telegram.RobToPlc.CyclicOptional.CartesianPosition.Turns_J6_J5          := RecvData.GetByte();
    Telegram.RobToPlc.CyclicOptional.CartesianPosition.Turns_E1             := RecvData.GetByte();
    Telegram.RobToPlc.CyclicOptional.CartesianPosition.E1                   := RecvData.GetReal();
    Telegram.RobToPlc.CyclicOptional.CartesianPosition.ToolNo               := RecvData.GetUsint();
    Telegram.RobToPlc.CyclicOptional.CartesianPosition.FrameNo              := RecvData.GetUsint();
    Telegram.RobToPlc.CyclicOptional.CartesianPosition.CurrentlyUsedToolNo  := RecvData.GetUsint();
    Telegram.RobToPlc.CyclicOptional.CartesianPosition.CurrentlyUsedFrameNo := RecvData.GetUsint();
    Telegram.RobToPlc.CyclicOptional.CartesianPosition.Reserve_1            := RecvData.GetByte();
    Telegram.RobToPlc.CyclicOptional.CartesianPosition.Reserve_2            := RecvData.GetByte();
  END_IF
  // }}}

  // AxesGroup.OptionalCyclic.RobToPlc.JointPosition {{{
  IF ( AxesGroup.CyclicOptional.RobToPlc.JointPosition.Active )
  THEN
    Telegram.RobToPlc.CyclicOptional.JointPosition.J1         := RecvData.GetReal();
    Telegram.RobToPlc.CyclicOptional.JointPosition.J2         := RecvData.GetReal();
    Telegram.RobToPlc.CyclicOptional.JointPosition.J3         := RecvData.GetReal();
    Telegram.RobToPlc.CyclicOptional.JointPosition.J4         := RecvData.GetReal();
    Telegram.RobToPlc.CyclicOptional.JointPosition.J5         := RecvData.GetReal();
    Telegram.RobToPlc.CyclicOptional.JointPosition.J6         := RecvData.GetReal();
    Telegram.RobToPlc.CyclicOptional.JointPosition.E1         := RecvData.GetReal();
    Telegram.RobToPlc.CyclicOptional.JointPosition.E1_Reserve := RecvData.GetWord();
  END_IF
  // }}}

  // AxesGroup.OptionalCyclic.RobToPlc.CartesianForce {{{
  IF ( AxesGroup.CyclicOptional.RobToPlc.Force.Active )
  THEN
    Telegram.RobToPlc.CyclicOptional.Force.X  := RecvData.GetReal();
    Telegram.RobToPlc.CyclicOptional.Force.Y  := RecvData.GetReal();
    Telegram.RobToPlc.CyclicOptional.Force.Z  := RecvData.GetReal();
    Telegram.RobToPlc.CyclicOptional.Force.Rx := RecvData.GetReal();
    Telegram.RobToPlc.CyclicOptional.Force.Ry := RecvData.GetReal();
    Telegram.RobToPlc.CyclicOptional.Force.Rz := RecvData.GetReal();
  END_IF
  // }}}

  // AxesGroup.OptionalCyclic.RobToPlc.Current {{{
  IF ( AxesGroup.CyclicOptional.RobToPlc.Current.Active )
  THEN
    Telegram.RobToPlc.CyclicOptional.Current.J1  := RecvData.GetReal();
    Telegram.RobToPlc.CyclicOptional.Current.J2  := RecvData.GetReal();
    Telegram.RobToPlc.CyclicOptional.Current.J3  := RecvData.GetReal();
    Telegram.RobToPlc.CyclicOptional.Current.J4  := RecvData.GetReal();
    Telegram.RobToPlc.CyclicOptional.Current.J5  := RecvData.GetReal();
    Telegram.RobToPlc.CyclicOptional.Current.J6  := RecvData.GetReal();
  END_IF

  // AxesGroup.OptionalCyclic.RobToPlc.CartesianPosExt {{{
  IF ( AxesGroup.CyclicOptional.RobToPlc.CartesianPositionExt.Active )
  THEN
    Telegram.RobToPlc.CyclicOptional.CartesianPositionExt.E2 := RecvData.GetReal();
    Telegram.RobToPlc.CyclicOptional.CartesianPositionExt.E3 := RecvData.GetReal();
    Telegram.RobToPlc.CyclicOptional.CartesianPositionExt.E4 := RecvData.GetReal();
    Telegram.RobToPlc.CyclicOptional.CartesianPositionExt.E5 := RecvData.GetReal();
    Telegram.RobToPlc.CyclicOptional.CartesianPositionExt.E6 := RecvData.GetReal();
  END_IF
  // }}}

  // AxesGroup.OptionalCyclic.RobToPlc.JointPosition {{{
  IF ( AxesGroup.CyclicOptional.RobToPlc.JointPositionExt.Active )
  THEN
    Telegram.RobToPlc.CyclicOptional.JointPositionExt.E2 := RecvData.GetReal();
    Telegram.RobToPlc.CyclicOptional.JointPositionExt.E3 := RecvData.GetReal();
    Telegram.RobToPlc.CyclicOptional.JointPositionExt.E4 := RecvData.GetReal();
    Telegram.RobToPlc.CyclicOptional.JointPositionExt.E5 := RecvData.GetReal();
    Telegram.RobToPlc.CyclicOptional.JointPositionExt.E6 := RecvData.GetReal();
  END_IF
  // }}}

  // AxesGroup.OptionalCyclic.RobToPlc.CartesianForceExt {{{
  IF ( AxesGroup.CyclicOptional.RobToPlc.ForceExt.Active )
  THEN
    Telegram.RobToPlc.CyclicOptional.ForceExt.E1  := RecvData.GetReal();
    Telegram.RobToPlc.CyclicOptional.ForceExt.E2  := RecvData.GetReal();
    Telegram.RobToPlc.CyclicOptional.ForceExt.E3  := RecvData.GetReal();
    Telegram.RobToPlc.CyclicOptional.ForceExt.E4  := RecvData.GetReal();
    Telegram.RobToPlc.CyclicOptional.ForceExt.E5  := RecvData.GetReal();
    Telegram.RobToPlc.CyclicOptional.ForceExt.E6  := RecvData.GetReal();
  END_IF
  // }}}

  // AxesGroup.OptionalCyclic.RobToPlc.CurrentExt {{{
  IF ( AxesGroup.CyclicOptional.RobToPlc.CurrentExt.Active )
  THEN
    Telegram.RobToPlc.CyclicOptional.CurrentExt.E1  := RecvData.GetReal();
    Telegram.RobToPlc.CyclicOptional.CurrentExt.E2  := RecvData.GetReal();
    Telegram.RobToPlc.CyclicOptional.CurrentExt.E3  := RecvData.GetReal();
    Telegram.RobToPlc.CyclicOptional.CurrentExt.E4  := RecvData.GetReal();
    Telegram.RobToPlc.CyclicOptional.CurrentExt.E5  := RecvData.GetReal();
    Telegram.RobToPlc.CyclicOptional.CurrentExt.E6  := RecvData.GetReal();
  END_IF
  // }}}

END_METHOD

METHOD PRIVATE ParseRecvPayloadFooter
VAR_IN_OUT
  /// Robot assignment of function
  AxesGroup : AxesGroup;
END_VAR

  Telegram.RobToPlc.Footer.LifeSign := RecvData.GetLifeSignFooter();

END_METHOD

METHOD PROTECTED ParseRecvPayloadHeader
VAR_IN_OUT
  /// Robot assignment of function
  AxesGroup    : AxesGroup;
END_VAR

  // Version
  Telegram.RobToPlc.Header.SRCIVersion := ByteToVersion(RecvData.GetByte());
  // Connection alive signal
  Telegram.RobToPlc.Header.LifeSign    := RecvData.GetHalfeByte2(IncPayloadPtr := TRUE);
  // Reserved byte
  Telegram.RobToPlc.Header.Reserved       := RecvData.GetByte();
  // Initialization and Telegram control state
  Telegram.RobToPlc.Header.TelegramState  := RecvData.GetUsint();
  // Combination of various RA related states.
  Telegram.RobToPlc.Header.StatusRobotArm := RecvData.GetDword();
  // Actual override in percentage encoding
  Telegram.RobToPlc.Header.Override       := RecvData.GetUint();

END_METHOD

METHOD PRIVATE ParseRecvPayloadLogging
VAR_IN_OUT
  /// Robot assignment of function
  AxesGroup    : AxesGroup;
END_VAR

VAR
  /// internal sequence index for loops
  _seqIdx : DINT;
  /// internal fragment index for loops
  _fragIdx : DINT;
END_VAR

  RETURN;
  FOR _seqIdx := 0 TO AxesGroup.State.SequenceCountRecv
  DO
    // check new data to receive ?
    IF ( Telegram.RobToPlc.Sequence[_seqIdx].Header.SEQ_ACK <> AxesGroup.State.LastACK[_seqIdx])
    THEN
      // Check sequence payload > 0 ?
      IF (Telegram.RobToPlc.Sequence[_seqIdx].Header.PayloadLength > 0)
      THEN
        // Create log entry
        CreateLogMessagePara4 ( Timestamp   := SystemTime,
                                MessageType := MessageType.CMD,
                                Severity    := Severity.DEBUG,
                                MessageCode := 0,
                                MessageText := 'RecvData: ACK = {1}, received Sequence [{2}] with PayloadLength = {3}, Lifesign = {4}',
                                Para1       :=  UINT_TO_STRING(Telegram.RobToPlc.Sequence[_seqIdx].Header.SEQ_ACK),
                                Para2       :=  DINT_TO_STRING(_seqIdx),
                                Para3       :=  UINT_TO_STRING(Telegram.RobToPlc.Sequence[_seqIdx].Header.PayloadLength),
                                Para4       :=  BYTE_TO_STRING(Telegram.RobToPlc.Header.LifeSign));

        FOR _fragIdx := 0 TO AxesGroup.State.FragmentCountRecv[_seqIdx]
        DO
          // Check fragment payload > 0 ?
          IF (Telegram.RobToPlc.Sequence[_seqIdx].Fragment[_fragIdx].Header.PayloadLength > 0)
          THEN
            // Create log entry
            CreateLogMessagePara5 ( Timestamp   := SystemTime,
                                    MessageType := MessageType.CMD,
                                    Severity    := Severity.DEBUG,
                                    MessageCode := 0,
                                    MessageText := 'RecvData: received Fragment [{1}] with PayloadLength = {2}, CmdID <{3}> , CmdState: {4}, Fragment-Action Bits: {5}',
                                    Para1       :=  DINT_TO_STRING(_fragIdx),
                                    Para2       :=  UINT_TO_STRING              (Telegram.RobToPlc.Sequence[_seqIdx].Fragment[_fragIdx].Header.PayloadLength),
                                    Para3       :=  DINT_TO_STRING              (Telegram.RobToPlc.Sequence[_seqIdx].Fragment[_fragIdx].Header.CmdID),
                                    Para4       :=  CMD_MESSAGE_STATE_TO_STRING (Telegram.RobToPlc.Sequence[_seqIdx].Fragment[_fragIdx].Command.Header.State),
                                    Para5       :=    FRAGMENT_ACTION_TO_STRING (Telegram.RobToPlc.Sequence[_seqIdx].Fragment[_fragIdx].Header.FragmentAction));
          END_IF
        END_FOR
      END_IF
    END_IF
  END_FOR

END_METHOD

METHOD PRIVATE ParseRecvPayloadSequence
VAR_IN_OUT
  /// Robot assignment of function
  AxesGroup        : AxesGroup;
END_VAR

VAR
  /// internal index
 _idx              : DINT;
  /// index for sequence
 _seqIdx           : DINT;
  /// index for fragment
 _fragIdx          : DINT;
  /// current payload pointer for current fragment
 _payLoadPtr       : DINT;
  /// Amount of sequences
 _seqCount         : DINT;
  /// current payload pointer of the current sequence
 _seqPayloadPtr    : UINT;
  /// ST-FIX F63: start of the payload of each sequence (behind its sequence header)
 _rcvStart         : ARRAY[0..1] OF DINT;
  /// ST-FIX F63: sequence that is processed first (lower Ack)
 _rcvFirst         : DINT;
  /// ST-FIX F63: loop counter over the sequences in Ack order
 _rcvOrderIdx      : DINT;
  /// ST-FIX F63: distance of the two Ack numbers
 _rcvDiff          : DINT;
END_VAR

  // Check 2nd sequence active ?
  IF ( _parCfg.Com.TwoSequences )
  THEN
   _seqCount := _seqCount + 1;
  END_IF

  // ST-FIX F63: read the headers of all sequences, each from its own address (Fig. 5-205)
  FOR _seqIdx := 0 TO _seqCount
  DO
    IF ( _seqIdx = PRIMARY_SEQUENCE )
    THEN
      RecvData.PayloadPtr := CalculateSequencePayloadStartAdr(AxesGroup := AxesGroup,
                                                              Direction := ComDirection.ROB_TO_PLC,
                                                              Sequence  := SequenceFlag.PRIMARY_SEQUENCE);
    ELSE
      RecvData.PayloadPtr := CalculateSequencePayloadStartAdr(AxesGroup := AxesGroup,
                                                              Direction := ComDirection.ROB_TO_PLC,
                                                              Sequence  := SequenceFlag.SECONDARY_SEQUENCE);
    END_IF

    // parse sequence header
    Telegram.RobToPlc.Sequence[_seqIdx].Header.SEQ_ACK       := RecvData.GetUint();
    Telegram.RobToPlc.Sequence[_seqIdx].Header.PayloadLength := RecvData.GetUint();
   _rcvStart[_seqIdx] := RecvData.PayloadPtr;
  END_FOR

  // ST-FIX F63: the sequence with the lower Ack first (Fig. 5-207/5-208), numbers wrap 254 -> 1
  _rcvFirst := 0;
  IF ( _seqCount = 1 )
  THEN
   _rcvDiff := UINT_TO_DINT(Telegram.RobToPlc.Sequence[0].Header.SEQ_ACK)
             - UINT_TO_DINT(Telegram.RobToPlc.Sequence[1].Header.SEQ_ACK);
    IF ( _rcvDiff < 0 ) THEN _rcvDiff := _rcvDiff + 254; END_IF
    IF (( _rcvDiff > 0 ) AND ( _rcvDiff < 127 )) THEN _rcvFirst := 1; END_IF
  END_IF

  FOR _rcvOrderIdx := 0 TO _seqCount
  DO
    IF ( _rcvOrderIdx = 0 ) THEN _seqIdx := _rcvFirst; ELSE _seqIdx := 1 - _rcvFirst; END_IF

    // ST-FIX F5: every sequence starts with fragment 0
    _fragIdx       := 0;
    _seqPayloadPtr := 0;
    RecvData.PayloadPtr := _rcvStart[_seqIdx];

    // check new data available ?
    // ST-FIX F63: only the Ack of the Seq that was sent (Seq = Ack) carries the response of it;
    // with two sequences the RC may send Ack 0 in the sequence it does not process
    IF (( Telegram.RobToPlc.Sequence[_seqIdx].Header.SEQ_ACK <> AxesGroup.State.LastACK[_seqIdx]    ) AND
        ( Telegram.RobToPlc.Sequence[_seqIdx].Header.SEQ_ACK  = AxesGroup.State.CurrentSEQ[_seqIdx] ))
    THEN
      // Check sequence payload available ?
      IF (Telegram.RobToPlc.Sequence[_seqIdx].Header.PayloadLength > 0)
      THEN
        // Check sequence payload length is valid ?
        IF ( Telegram.RobToPlc.Sequence[_seqIdx].Header.PayloadLength > _parCfg.Com.TelegramLengthRobToPlc )
        THEN
          // Create log entry for payload not valid
          CreateLogMessagePara2 ( Timestamp   := SystemTime,
                                  MessageType := MessageType.CMD,
                                  Severity    := Severity.DEBUG,
                                  MessageCode := 0,
                                  MessageText := 'Invalid sequence payload length, Sequence = {1}, PayloadLength = {2} ',
                                  Para1       :=  DINT_TO_STRING(_seqIdx),
                                  Para2       :=  UINT_TO_STRING(Telegram.RobToPlc.Sequence[_seqIdx].Header.PayloadLength));
                                  RETURN;
        ELSE
          // Create log entry
          CreateLogMessagePara4 ( Timestamp   := SystemTime,
                                  MessageType := MessageType.CMD,
                                  Severity    := Severity.DEBUG,
                                  MessageCode := 0,
                                  MessageText := 'RecvData: ACK = {1}, received Sequence [{2}] with PayloadLength = {3}, Lifesign = {4}',
                                  Para1       :=  UINT_TO_STRING(Telegram.RobToPlc.Sequence[_seqIdx].Header.SEQ_ACK),
                                  Para2       :=  DINT_TO_STRING(_seqIdx),
                                  Para3       :=  UINT_TO_STRING(Telegram.RobToPlc.Sequence[_seqIdx].Header.PayloadLength),
                                  Para4       :=  BYTE_TO_STRING(Telegram.RobToPlc.Header.LifeSign));
        END_IF

        // processing sequence payload
        WHILE ( _seqPayloadPtr < Telegram.RobToPlc.Sequence[_seqIdx].Header.PayloadLength )
        DO
          // parse header
          Telegram.RobToPlc.Sequence[_seqIdx].Fragment[_fragIdx].Header.CmdID          := RecvData.GetUint();
          Telegram.RobToPlc.Sequence[_seqIdx].Fragment[_fragIdx].Header.Reserve        := RecvData.GetByte();
          Telegram.RobToPlc.Sequence[_seqIdx].Fragment[_fragIdx].Header.FragmentAction := RecvData.GetByte();
          Telegram.RobToPlc.Sequence[_seqIdx].Fragment[_fragIdx].Header.PayloadPointer := RecvData.GetUint();
          Telegram.RobToPlc.Sequence[_seqIdx].Fragment[_fragIdx].Header.PayloadLength  := RecvData.GetUint();

          // add header size to payload pointer
         _seqPayloadPtr := _seqPayloadPtr + SIZEOF(Telegram.RobToPlc.Sequence[_seqIdx].Fragment[_fragIdx].Header);

          // Check fragment payload available ?
          IF (Telegram.RobToPlc.Sequence[_seqIdx].Fragment[_fragIdx].Header.PayloadLength > 0)
          THEN
            // Check fragment payload length is valid ?
            IF ( Telegram.RobToPlc.Sequence[_seqIdx].Fragment[_fragIdx].Header.PayloadLength > _parCfg.Com.TelegramLengthRobToPlc )
            THEN
              // Create log entry for payload not valid
              CreateLogMessagePara2 ( Timestamp   := SystemTime,
                                      MessageType := MessageType.CMD,
                                      Severity    := Severity.DEBUG,
                                      MessageCode := 0,
                                      MessageText := 'Invalid fragment payload length, Sequence = {1}, PayloadLength = {2} ',
                                      Para1       :=  DINT_TO_STRING(_seqIdx),
                                      Para2       :=  UINT_TO_STRING(Telegram.RobToPlc.Sequence[_seqIdx].Fragment[_fragIdx].Header.PayloadLength));
                                      RETURN;
            END_IF

            // Fill Response payload
            FOR _idx := 0 TO Telegram.RobToPlc.Sequence[_seqIdx].Fragment[_fragIdx].Header.PayloadLength -1
            DO
              // calculate payload pointer
             _payLoadPtr := Telegram.RobToPlc.Sequence[_seqIdx].Fragment[_fragIdx].Header.PayloadPointer + _idx;

              IF (( _payLoadPtr >= 0                                          ) AND
                  ( _payLoadPtr <= RobotLibraryParameter.RESPONSE_PAYLOAD_MAX ))
              THEN
                Telegram.RobToPlc.Sequence[_seqIdx].Fragment[_fragIdx].Command.Payload[_payLoadPtr] := RecvData.GetByte();
                // inc payload pointer
               _seqPayloadPtr := _seqPayloadPtr + SIZEOF(BYTE);
              ELSE
                // Create log entry for payload pointer not valid
                CreateLogMessagePara3 ( Timestamp   := SystemTime,
                                        MessageType := MessageType.CMD,
                                        Severity    := Severity.DEBUG,
                                        MessageCode := 0,
                                        MessageText := 'Invalid fragment payload pointer, Sequence = {1}, Fragment = {2}, PayloadPointer = {3} ',
                                        Para1       :=  DINT_TO_STRING(_seqIdx),
                                        Para2       :=  DINT_TO_STRING(_fragIdx),
                                        Para3       :=  DINT_TO_STRING(_payLoadPtr));
                                        RETURN;
  					  END_IF

            END_FOR

            // Add Response to ACR
            AxesGroup.Acyclic.ActiveCommandRegister.AddRsp(Telegram.RobToPlc.Sequence[_seqIdx].Fragment[_fragIdx]);

            // Only for debugging - header is part of the payload itself
            Telegram.RobToPlc.Sequence[_seqIdx].Fragment[_fragIdx].Command.Header.State                 :=      GetHalfeByteLo( Value :=  Telegram.RobToPlc.Sequence[_seqIdx].Fragment[_fragIdx].Command.Payload[0]);
            Telegram.RobToPlc.Sequence[_seqIdx].Fragment[_fragIdx].Command.Header.ParSeq                :=      GetHalfeByteHi( Value :=  Telegram.RobToPlc.Sequence[_seqIdx].Fragment[_fragIdx].Command.Payload[0]);
            Telegram.RobToPlc.Sequence[_seqIdx].Fragment[_fragIdx].Command.Header.AlarmMessageSeverity  :=        BYTE_TO_SINT(           Telegram.RobToPlc.Sequence[_seqIdx].Fragment[_fragIdx].Command.Payload[1]);
            Telegram.RobToPlc.Sequence[_seqIdx].Fragment[_fragIdx].Command.Header.AlarmMessageCode      :=  CombineBytesToUint( HiByte := Telegram.RobToPlc.Sequence[_seqIdx].Fragment[_fragIdx].Command.Payload[2],
                                                                                                                                LoByte := Telegram.RobToPlc.Sequence[_seqIdx].Fragment[_fragIdx].Command.Payload[3]);
            // Create log entry
            CreateLogMessagePara5 ( Timestamp   := SystemTime,
                                    MessageType := MessageType.CMD,
                                    Severity    := Severity.DEBUG,
                                    MessageCode := 0,
                                    MessageText := 'RecvData: received Fragment [{1}] with PayloadLength = {2}, CmdID <{3}> , CmdState: {4}, Fragment-Action Bits: {5}',
                                    Para1       :=  DINT_TO_STRING(_seqIdx),
                                    Para2       :=  UINT_TO_STRING              (Telegram.RobToPlc.Sequence[_seqIdx].Fragment[_fragIdx].Header.PayloadLength),
                                    Para3       :=  DINT_TO_STRING              (Telegram.RobToPlc.Sequence[_seqIdx].Fragment[_fragIdx].Header.CmdID),
                                    Para4       :=  CMD_MESSAGE_STATE_TO_STRING (Telegram.RobToPlc.Sequence[_seqIdx].Fragment[_fragIdx].Command.Header.State),
                                    Para5       :=    FRAGMENT_ACTION_TO_STRING (Telegram.RobToPlc.Sequence[_seqIdx].Fragment[_fragIdx].Header.FragmentAction));
          END_IF

          // Check still payload left ? -> goto next fragment
          IF ( _seqPayloadPtr < Telegram.RobToPlc.Sequence[_seqIdx].Header.PayloadLength )
          THEN
           _fragIdx := _fragIdx + 1;
          END_IF

          // Check fragment index limit reached ?
          IF ( _fragIdx > RobotLibraryParameter.FRAGMENT_MAX )
          THEN
            // Create log entry
            CreateLogMessagePara1 ( Timestamp   := SystemTime,
                                    MessageType := MessageType.CMD,
                                    Severity    := Severity.ERROR, // ST-FIX F52: responses are lost
                                    MessageCode := 0,
                                    MessageText := 'Fragment index out of range, _fragIdx = {1} ',
                                    Para1       :=  DINT_TO_STRING(_fragIdx));
                                    RETURN;
          END_IF
        END_WHILE
      END_IF
    END_IF
  END_FOR

END_METHOD

METHOD Reset
VAR_IN_OUT
  /// Robot assignment of function
  AxesGroup : AxesGroup;
END_VAR

  // reset flags
  Busy              := FALSE;
  Initialized       := FALSE;
  Synchronized      := FALSE;
  Error             := FALSE;
  ErrorID           := 0;
  ErrorAddTxt       := '';
  WarningID         := 0;
  InfoID            := 0;

  // Reset internal functon blocks
  _exchangeConfiguration      .Enable  := FALSE;
  _readRobotData              .Execute := FALSE;
  _readMessages               .Enable  := FALSE;
  _readToolData               .Execute := FALSE;
  _readFrameData              .Execute := FALSE;
  _readLoadData               .Execute := FALSE;
  _readWorkArea               .Execute := FALSE;
  _readRobotSWLimits          .Execute := FALSE;
  _readRobotDefaultDynamics   .Execute := FALSE;
  _readRobotReferenceDynamics .Execute := FALSE;
  _writeToolData              .Execute := FALSE;
  _writeFrameData             .Execute := FALSE;
  _writeLoadData              .Execute := FALSE;
  _writeWorkArea              .Execute := FALSE;
  _writeRobotSWLimits         .Execute := FALSE;
  _writeRobotDefaultDynamics  .Execute := FALSE;
  _writeRobotReferenceDynamics.Execute := FALSE;

  // Set Client error to force server error
  AxesGroup.Cyclic.PlcToRob.Control := ControlHalfByte.NONE;

  // Reset synchronisation state variables
  AxesGroup.State.SyncStatePlc.InSync.Frame             := FALSE;
  AxesGroup.State.SyncStatePlc.InSync.Tool              := FALSE;
  AxesGroup.State.SyncStatePlc.InSync.Load              := FALSE;
  AxesGroup.State.SyncStatePlc.InSync.WorkArea          := FALSE;
  AxesGroup.State.SyncStatePlc.InSync.SwLimits          := FALSE;
  AxesGroup.State.SyncStatePlc.InSync.DefaultDynamics   := FALSE;
  AxesGroup.State.SyncStatePlc.InSync.ReferenceDynamics := FALSE;

  AxesGroup.State.SyncStatePlc.UnSyncNo.Frame    := 0;
  AxesGroup.State.SyncStatePlc.UnSyncNo.Tool     := 0;
  AxesGroup.State.SyncStatePlc.UnSyncNo.Load     := 0;
  AxesGroup.State.SyncStatePlc.UnSyncNo.WorkArea := 0;

  AxesGroup.State.SyncStateRc .InSync.Frame             := FALSE;
  AxesGroup.State.SyncStateRc .InSync.Tool              := FALSE;
  AxesGroup.State.SyncStateRc .InSync.Load              := FALSE;
  AxesGroup.State.SyncStateRc .InSync.WorkArea          := FALSE;
  AxesGroup.State.SyncStateRc .InSync.SwLimits          := FALSE;
  AxesGroup.State.SyncStateRc .InSync.DefaultDynamics   := FALSE;
  AxesGroup.State.SyncStateRc .InSync.ReferenceDynamics := FALSE;

  AxesGroup.State.SyncStateRc .UnSyncNo.Frame    := 0;
  AxesGroup.State.SyncStateRc .UnSyncNo.Tool     := 0;
  AxesGroup.State.SyncStateRc .UnSyncNo.Load     := 0;
  AxesGroup.State.SyncStateRc .UnSyncNo.WorkArea := 0;

  // Reset active command register
  AxesGroup.Acyclic.ActiveCommandRegister.Reset();

  // reset step counters
  _stepCmd                   := 0;
  _stepSyncFrameData         := 0;
  _stepSyncLoadData          := 0;
  _stepSyncDefaultDynamics   := 0;
  _stepSyncReferenceDynamics := 0;
  _stepSyncSWLimits          := 0;
  _stepSyncToolData          := 0;
  _stepSyncWorkArea          := 0;

END_METHOD

METHOD PUBLIC SetError
VAR_INPUT
  /// ErrorID reported by RC for error identification according to Table 7-1
  ErrorID   : WORD;
  /// TRUE = overwrite an existing error
  Overwrite : BOOL;
END_VAR

  IF ( NOT HasError ) OR ( Overwrite )
  THEN
    THIS^.ErrorID := ErrorID;
  END_IF

END_METHOD

METHOD PUBLIC SetInfo
VAR_INPUT
  /// InfoID for info identification reported during execution of command according to Table 7-5
  InfoID    : WORD;
  /// TRUE = overwrite an existing info
  Overwrite : BOOL;
END_VAR

  IF ( NOT HasInfo ) OR ( Overwrite )
  THEN
    THIS^.InfoID := InfoID;
  END_IF

END_METHOD

METHOD PUBLIC SetWarning
VAR_INPUT
  /// WarningID for warning identification reported during execution of command according to Table 7-3
  WarningID : WORD;
  /// TRUE = overwrite an existing warning
  Overwrite : BOOL;
END_VAR

  IF ( NOT HasWarning ) OR ( Overwrite )
  THEN
    THIS^.WarningID := WarningID;
  END_IF

END_METHOD

/// ST-FIX F130: TRUE when the synchronization modes of a data set are defined
/// (during the start-up NO_SYNCHRONIZATION .. SERVER_TO_CLIENT, after the start-up also AUTOMATIC)
METHOD PRIVATE SyncModesValid : BOOL
VAR_INPUT
  /// Synchronization mode during the start-up
  During : SyncMode;
  /// Synchronization mode after the start-up
  After  : SyncMode;
END_VAR

  SyncModesValid := ( During >= SyncMode.NO_SYNCHRONIZATION ) AND
                    ( During <  SyncMode.AUTOMATIC          ) AND
                    ( After  >= SyncMode.NO_SYNCHRONIZATION ) AND
                    ( After  <= SyncMode.AUTOMATIC          );

END_METHOD
